Fanuc KAREL source: KD00067.KL

PROGRAM KD00067
%NOLOCKGROUP
VAR
  I: INTEGER
  J: INTEGER
  B: BOOLEAN
  R: REAL
  S: STRING[80]
BEGIN
  CONDITION[1]:
  WHEN DIN[1] = ON DO
    PAUSE
  ENDCONDITION
END KD00067
